(* IEC 61131-3 sources: plcassist-cli/packages/volt-lsp-iec/test-corpus/pro2193/Device/Plc Logic/Application/99 Library/Function Blocks/Actuators/Conveyors, 3 files *)

(* ---- ConveyorAdjustableSpeedFB.fb ---- *)
{attribute 'symbol' := 'none'}
FUNCTION_BLOCK PUBLIC ConveyorAdjustableSpeedFB
EXTENDS ConveyorFB
IMPLEMENTS IActuator
VAR_INPUT
	xAutoCycleActive	: BOOL;
END_VAR
VAR CONSTANT
	rMaxSpeedSetting	: REAL	:= 150.0;	// Upper limit of speed setpoint (in Hz). Set limit for rSetPointSpeed value in HMI.
END_VAR

SUPER^(profile := profile);

END_FUNCTION_BLOCK

// Maps the actuator to the physical output
METHOD MapAnalogOut : WORD
IF xAutoCycleActive OR Output.Map() THEN
	MapAnalogOut	:= RANGE_TO_WORD(input := profile.rVel, input_LO := 0.0, input_HI := rMaxSpeedSetting);
ELSE
	MapAnalogOut	:= WORD#0;
END_IF
END_METHOD

(* ---- ConveyorFB.fb ---- *)
{attribute 'symbol' := 'none'}
FUNCTION_BLOCK PUBLIC ConveyorFB
EXTENDS ActuatorWithManualControlAndAlarm_BaseFB
IMPLEMENTS IActuator
VAR_INPUT
	{attribute 'symbol' := 'read'}	beltRunning				: BOOL;
	errorId					: WORD;
END_VAR
VAR_IN_OUT
	profile					: ProfileType;
END_VAR
VAR
	NotRunningAlarm			: SetErrorFB;
	{attribute 'symbol' := 'read'}	Output					: ActuatorFB;
	beltStarted				: BTON;
	beltStopped				: BTOF;
END_VAR

SUPER^();

// Instantiate the output
Output();

UpdateTimers();

END_FUNCTION_BLOCK

METHOD PROTECTED Alarms
NotRunningAlarm(
	moduleHandler	:= moduleHandler,
	textRefId		:= textRefId,
	alarmCondition	:= alarmEnable AND (beltRunning XOR Output.Map()),
	alarmDelay		:= alarmDelay,
	errorId			:= errorId,
	severity		:= severity,
	reaction		:= reaction,
	active			=> );
END_METHOD

METHOD PROTECTED ManualControl
VAR_INPUT
	minButtonPushed			: BOOL;		// Both the software button (on screen) and the hardware button (if attached)
	plusButtonPushed		: BOOL;		// Both the software button (on screen) and the hardware button (if attached)
END_VAR
IF plusButtonPushed THEN
	Set();
END_IF

IF minButtonPushed THEN
	Reset();
END_IF
END_METHOD

// Maps the actuator to the physical output
METHOD Map : BOOL
Map := Output.Map();
END_METHOD

// Reset the output (=False)
METHOD Reset
Output.Reset();

UpdateTimers();
END_METHOD

// Set the output (=True)
METHOD Set : BOOL
Output.Set();

UpdateTimers();
END_METHOD

// Set the output True or False
METHOD SetOrReset
VAR_INPUT
	xValue	: BOOL;
END_VAR
Output.SetOrReset(xValue);

UpdateTimers();
END_METHOD

METHOD PRIVATE UpdateTimers
beltStarted.Set(Output.Map(), profile.rAcc);
beltStopped.Set(Output.Map(), profile.rDec);
END_METHOD

{attribute 'monitoring':='call'}
PROPERTY PUBLIC ConveyorState : enumConveyorRunning_State
GET
VAR
END_VAR
IF NOT beltStopped.Q THEN
	ConveyorState	:= enumConveyorRunning_State.Standstill;
ELSIF beltStarted.Q THEN
	ConveyorState	:= enumConveyorRunning_State.ConstantVelocity;
ELSIF Output.Map() THEN
	ConveyorState	:= enumConveyorRunning_State.Accelerating;
ELSE
	ConveyorState	:= enumConveyorRunning_State.Decelerating;
END_IF
END_GET
END_PROPERTY

(* ---- ConveyorReversibleFB.fb ---- *)
{attribute 'symbol' := 'none'}
FUNCTION_BLOCK PUBLIC ConveyorReversibleFB
EXTENDS ConveyorFB
IMPLEMENTS IActuator
VAR
	{attribute 'symbol' := 'read'}	OutputReverse			: ActuatorFB;
END_VAR

SUPER^(profile := profile);

// Instantiate the output
OutputReverse();

END_FUNCTION_BLOCK

METHOD PROTECTED Alarms
NotRunningAlarm(
	moduleHandler	:= moduleHandler,
	textRefId		:= textRefId,
	alarmCondition	:= alarmEnable AND (beltRunning XOR (Output.Map() OR OutputReverse.Map())),
	alarmDelay		:= alarmDelay,
	errorId			:= errorId,
	severity		:= severity,
	reaction		:= reaction,
	active			=> );
END_METHOD

METHOD PROTECTED ManualControl
VAR_INPUT
	minButtonPushed			: BOOL;		// Both the software button (on screen) and the hardware button (if attached)
	plusButtonPushed		: BOOL;		// Both the software button (on screen) and the hardware button (if attached)
END_VAR
IF plusButtonPushed THEN
	IF Output.Map() THEN	// Conveyor moving forward
		Reset();
	ELSE
		Set();
	END_IF
END_IF

IF minButtonPushed THEN
	IF OutputReverse.Map() THEN	// Conveyor moving in reverse
		Reset();
	ELSE
		Reverse();
	END_IF
END_IF
END_METHOD

// Maps the actuator to start conveyor in reverse
METHOD MapReverse : BOOL
MapReverse := OutputReverse.Map();
END_METHOD

// Reset the output (=False)
METHOD Reset
SUPER^.Reset();
OutputReverse.Reset();
END_METHOD

METHOD Reverse : BOOL
VAR_INPUT
END_VAR
SUPER^.Set();
OutputReverse.Set();
END_METHOD

// Set the output (=True)
METHOD Set : BOOL
SUPER^.Set();
OutputReverse.Reset();
END_METHOD
